FUNCTION_BLOCK EEE_Bruto_HMI (* Service Interface Function Block Type *)
  (* Standard: 61499-2 *)
  (* Version 1.3, 21/10/2026, Hidryco, Hidryco, IHM da EEE_Bruto 1.3: ajustes nos sub-CATs Necessidade/Revezamento/PID; reset cmdResetFalhas / E_RESET_FALHAS_PROCESSO (legado) *)
  PACKAGE Hidryco.HidrycoLib;
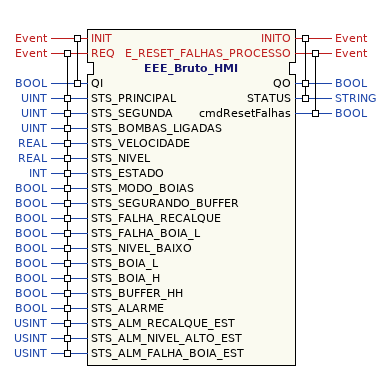
  EVENT_INPUT
    INIT WITH QI;
    REQ WITH STS_PRINCIPAL, STS_SEGUNDA, STS_BOMBAS_LIGADAS, STS_VELOCIDADE, STS_NIVEL, STS_ESTADO, STS_MODO_BOIAS, STS_SEGURANDO_BUFFER, STS_FALHA_RECALQUE, STS_FALHA_BOIA_L, STS_NIVEL_BAIXO, STS_BOIA_L, STS_BOIA_H, STS_BUFFER_HH, STS_ALARME, STS_ALM_RECALQUE_EST, STS_ALM_NIVEL_ALTO_EST, STS_ALM_FALHA_BOIA_EST; (* Atualizacao de status *)
  END_EVENT
  EVENT_OUTPUT
    INITO WITH QO, STATUS;
    E_RESET_FALHAS_PROCESSO WITH cmdResetFalhas;
  END_EVENT
  VAR_INPUT
    QI : BOOL;
    STS_PRINCIPAL : UINT; (* Bomba principal *)
    STS_SEGUNDA : UINT; (* Bomba que entra como 2a *)
    STS_BOMBAS_LIGADAS : UINT; (* Bombas ligadas *)
    STS_VELOCIDADE : REAL; (* Velocidade enviada as bombas (Hz) *)
    STS_NIVEL : REAL; (* Nivel do poco (LIT-03) *)
    STS_ESTADO : INT; (* 0 parada, 1 bombeando, 2 segurando (HH Nereda), 3 pelas boias, 4 falha de recalque, 5 nivel baixo (LSL), 6 automatico desabilitado, 7 emergencia *)
    STS_MODO_BOIAS : BOOL; (* Operacao pelas boias (LIT-03 em falha) *)
    STS_SEGURANDO_BUFFER : BOOL; (* Segurando o esgoto (HH do tanque do Nereda) *)
    STS_FALHA_RECALQUE : BOOL; (* Falha de recalque *)
    STS_FALHA_BOIA_L : BOOL; (* Boia LSL com defeito *)
    STS_NIVEL_BAIXO : BOOL; (* LSL abaixada: bombas intertravadas *)
    STS_BOIA_L : BOOL; (* LSL-04 levantada *)
    STS_BOIA_H : BOOL; (* LSH-05 levantada *)
    STS_BUFFER_HH : BOOL; (* HH do tanque do Nereda *)
    STS_ALARME : BOOL; (* Algum alarme da elevatoria *)
    STS_ALM_RECALQUE_EST : USINT; (* Estado do ALARM_BIT falha de recalque (0 normal, 1 ativo reconhecido, 2 ativo nao reconhecido, 3 saiu nao reconhecido, 4 ativo e saiu nao reconhecido) *)
    STS_ALM_NIVEL_ALTO_EST : USINT; (* Estado do ALARM_BIT nivel alto (LSH) (0 normal, 1 ativo reconhecido, 2 ativo nao reconhecido, 3 saiu nao reconhecido, 4 ativo e saiu nao reconhecido) *)
    STS_ALM_FALHA_BOIA_EST : USINT; (* Estado do ALARM_BIT defeito da boia LSL (0 normal, 1 ativo reconhecido, 2 ativo nao reconhecido, 3 saiu nao reconhecido, 4 ativo e saiu nao reconhecido) *)
  END_VAR
  VAR_OUTPUT
    QO : BOOL; (* Event Output Qualifier *)
    STATUS : STRING; (* Service Status *)
    cmdResetFalhas : BOOL; (* Reset das falhas da elevatoria (recalque, boia) e reconhecimento *)
  END_VAR
  SERVICE /
    SEQUENCE 
    END_SEQUENCE
  END_SERVICE
END_FUNCTION_BLOCK
